Fanuc KAREL source: kt00074.KL

-- PROVISIONAL review KL for V940-1; original PC SHA256 1a235635930bd4a78c076a49aaa3d7ae622327e0b629aee441ee8b36bd26a39a
-- Incomplete behavior may be omitted. Consult companion uncertainty JSON. Do not deploy.
PROGRAM KT00074
%NOLOCKGROUP
VAR
  R1 : REAL
  I2 : INTEGER
  OUT : REAL
BEGIN
  -- V9_ZERO_TABLE_METADATA_HINT layout=0001; no indexed target words; source/name/runtime held
  -- UNRESOLVED_PC offsets 5-16; opcodes 2E,23
  -- UNRESOLVED_PC offsets 21-32; opcodes 2E,23
  -- UNRESOLVED_PC offsets 37-57; opcodes 21,21,64,6B,23
  -- UNRESOLVED_PC offsets 62-66; opcodes 7F
END KT00074
